Fanuc KAREL source: kc00032.KL

-- PROVISIONAL review KL for V940-1; original PC SHA256 55ad30ce2591bec7ca28b17a5df9bf37aa6f2813eba171134a4edb4d7b463b68
-- Incomplete behavior may be omitted. Consult companion uncertainty JSON. Do not deploy.
PROGRAM KC00032
%NOLOCKGROUP
BEGIN
  -- V9_ZERO_TABLE_METADATA_HINT layout=0002_ascii; no indexed target words; source/name/runtime held
  -- UNRESOLVED_PC offsets 5-55; opcodes 27,22,2A,22,22,22,22,22,22,27,9D,31
  -- UNRESOLVED_PC offsets 60-64; opcodes 7F
END KC00032
